// SIMATIC S7-200 project (STEP 7-Micro/WIN), CPU 214 REL 00.91

SYMBOL_TABLE USUARIO1
IGNICION         Q0.5     //  RELE QUE PUENTEA EL TT DE HONEYWEEL
CALOR            I0.3     // SOLICITUD DE LLAMA POR FY800
APG              M0.0     // POSTPURGA DE APAGADOR
HW               Q0.4     // ENCENDIDO DEL HONEYWELL
M2               Q0.3     // CONTACTOR C1
M1D              Q0.2     // CONTACTOR DELTA
M1E              Q0.1     // CONTACTOR DE ARRANQUE ESTRELLA
M1P              Q0.0     // CONTACTOR PRICIPAL DE ARRANQUE ESTRELLA DELTA
STP              I0.1     // STOP DEL PROGRAMA
P_EMERG          I0.2     // PARO DE EMERGENCIA
START            I0.0     // INICIO DEL PROGRAMA
END_SYMBOL_TABLE

ORGANIZATION_BLOCK PRINCIPAL:OB1
TITLE=COMENTARIOS DEL PROGRAMA
BEGIN
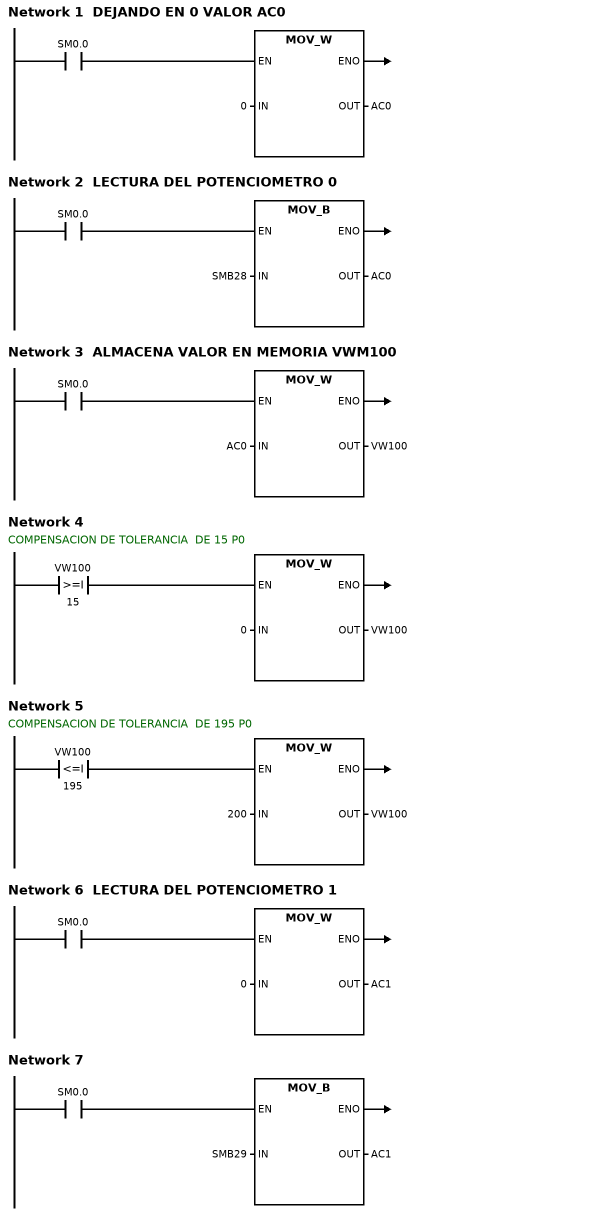
Network 1 // DEJANDO EN 0 VALOR AC0 
LD     SM0.0
MOVW   0, AC0
Network 2 // LECTURA DEL POTENCIOMETRO 0
// (network saved uncompiled; LAD cells follow)
// row 0: c0 -| |- SM0.0  c1 --  c2 [MOV_B EN:=power@row0, IN:=SMB28, ENO=>power, OUT=>AC0]  c3 ->
// row 1: c2 [box]
Network 3 // ALMACENA VALOR EN MEMORIA VWM100
LD     SM0.0
MOVW   AC0, VW100
Network 4
// COMPENSACION DE TOLERANCIA  DE 15 P0
LDW>=  VW100, 15
MOVW   0, VW100
Network 5
// COMPENSACION DE TOLERANCIA  DE 195 P0
LDW<=  VW100, 195
MOVW   200, VW100
Network 6 // LECTURA DEL POTENCIOMETRO 1
LD     SM0.0
MOVW   0, AC1
Network 7
LD     SM0.0
MOVB   SMB29, AC1
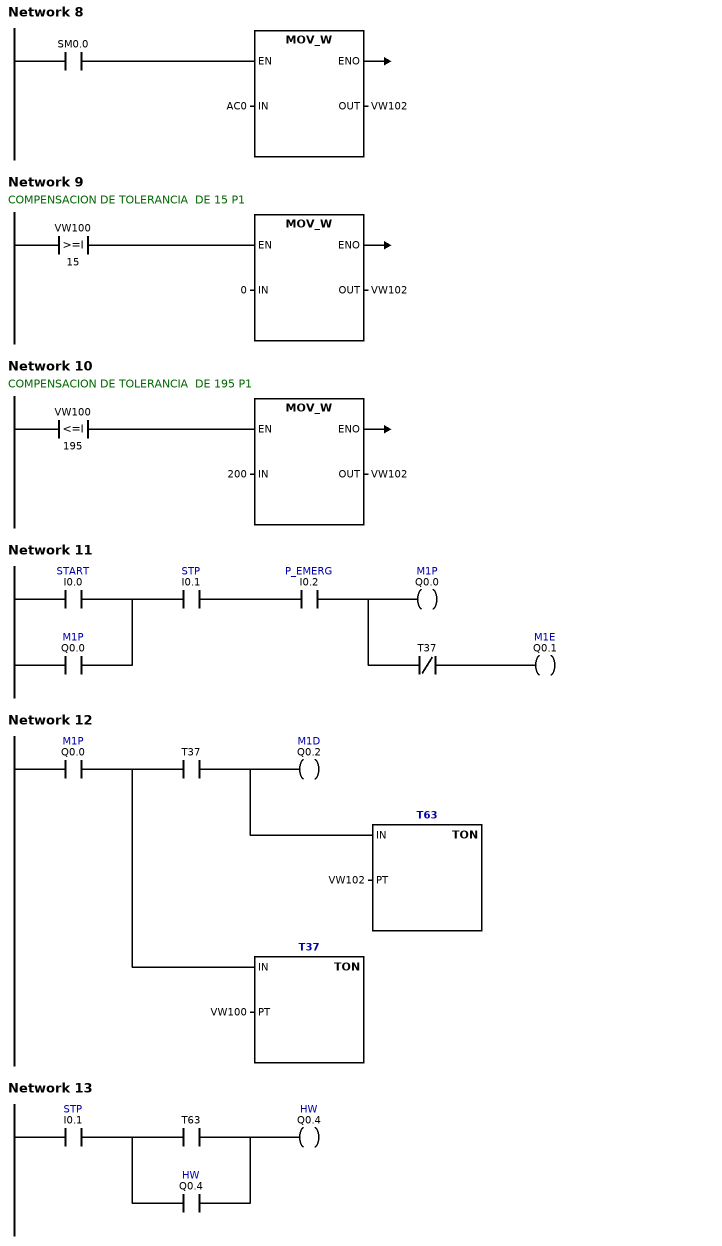
Network 8
LD     SM0.0
MOVW   AC0, VW102
Network 9
// COMPENSACION DE TOLERANCIA  DE 15 P1
LDW>=  VW100, 15
MOVW   0, VW102
Network 10
// COMPENSACION DE TOLERANCIA  DE 195 P1
LDW<=  VW100, 195
MOVW   200, VW102
Network 11
LD     START:I0.0
O      M1P:Q0.0
A      STP:I0.1
A      P_EMERG:I0.2
=      M1P:Q0.0
AN     T37
=      M1E:Q0.1
Network 12
LD     M1P:Q0.0
LPS
A      T37
=      M1D:Q0.2
TON    T63, VW102
LPP
TON    T37, VW100
Network 13
LD     STP:I0.1
LD     T63
O      HW:Q0.4
ALD
=      HW:Q0.4
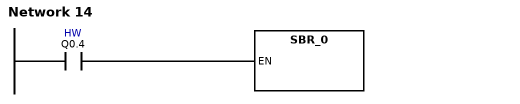
Network 14
LD     HW:Q0.4
CALL   SBR_0:SBR0
END_ORGANIZATION_BLOCK

SUBROUTINE_BLOCK SBR_0:SBR0
TITLE=COMENTARIOS DE LA SUBRUTINA
BEGIN
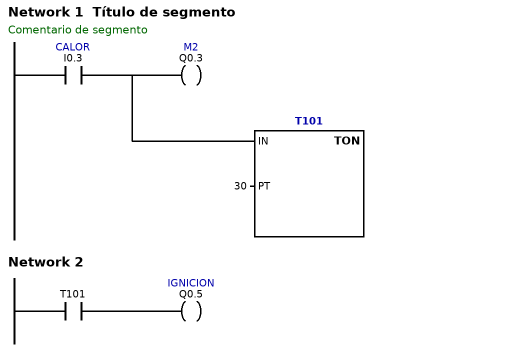
Network 1 // Título de segmento
// Comentario de segmento
LD     CALOR:I0.3
=      M2:Q0.3
TON    T101, 30
Network 2
LD     T101
=      IGNICION:Q0.5
END_SUBROUTINE_BLOCK
